PROGRAM PRG_IO_In
VAR
    fbSimInfeed, fbSimOutfeed, fbSimEjector, fbSimClamp, fbSimDiverter : FB_CylinderSim;
    fbSimCW : FB_CwSim;
END_VAR

IF GVL_Ctrl.xSim THEN
    //================ SIMULATION =================
    fbSimInfeed(  xValveWork := GVL_IO.stInfeed.xValveWork,   xValveHome := GVL_IO.stInfeed.xValveHome,
                  xSensWork => GVL_IO.stInfeed.xSensWork,     xSensHome => GVL_IO.stInfeed.xSensHome);
    fbSimOutfeed( xValveWork := GVL_IO.stOutfeed.xValveWork,  xValveHome := GVL_IO.stOutfeed.xValveHome,
                  xSensWork => GVL_IO.stOutfeed.xSensWork,    xSensHome => GVL_IO.stOutfeed.xSensHome);
    fbSimEjector( xValveWork := GVL_IO.stEjector.xValveWork,  xValveHome := GVL_IO.stEjector.xValveHome,
                  xSensWork => GVL_IO.stEjector.xSensWork,    xSensHome => GVL_IO.stEjector.xSensHome);
    fbSimClamp(   xValveWork := GVL_IO.stClamp.xValveWork,    xValveHome := GVL_IO.stClamp.xValveHome,
                  xSensWork => GVL_IO.stClamp.xSensWork,      xSensHome => GVL_IO.stClamp.xSensHome);
    fbSimDiverter(xValveWork := GVL_IO.stDiverter.xValveWork, xValveHome := GVL_IO.stDiverter.xValveHome,
                  xSensWork => GVL_IO.stDiverter.xSensWork,   xSensHome => GVL_IO.stDiverter.xSensHome);

    fbSimCW(xEnable := GVL_IO.xLaserEnable AND GVL_IO.xCW_STO,
            xTrig   := GVL_IO.xCW_Trig,
            nJob    := GVL_IO.nCW_Job,
            xReady  => GVL_IO.xCW_Lready,
            xJobLoaded => GVL_IO.xCW_JobLoaded,
            xBusy   => GVL_IO.xCW_MarkBusy);

    // part leaves the infeed barrier when the infeed cylinder pushed it;
    // part appears at the outfeed barrier after the ejector pushed a GOOD part (no bypass),
    // and disappears when the outfeed cylinder took it.
    IF GVL_IO.stInfeed.xSensWork THEN
        GVL_Ctrl.xSimPartIn := FALSE;
    END_IF
    IF GVL_IO.stEjector.xSensWork AND NOT GVL_IO.xBypassAS THEN
        GVL_Ctrl.xSimPartOut := TRUE;
    ELSIF GVL_IO.stOutfeed.xSensWork THEN
        GVL_Ctrl.xSimPartOut := FALSE;
    END_IF

    GVL_IO.xEStop          := GVL_Ctrl.xSimEStop;
    GVL_IO.xPressureOK     := GVL_Ctrl.xSimPressureOK;
    GVL_IO.xLS_Infeed      := GVL_Ctrl.xSimPartIn;
    GVL_IO.xLS_Outfeed     := GVL_Ctrl.xSimPartOut;
    GVL_IO.xServoInLatched := TRUE;   GVL_IO.xServoInAS  := FALSE;  GVL_IO.xServoInGS  := TRUE;
    GVL_IO.xServoOutLatched:= TRUE;   GVL_IO.xServoOutAS := FALSE;  GVL_IO.xServoOutGS := TRUE;
ELSE
    //================ REAL HARDWARE =================
    GVL_IO.xPressureOK     := GVL_HW.xMaintPressureOK;
    GVL_IO.xEStop          := GVL_HW.xEStopPressed;
    GVL_IO.xLS_Infeed      := GVL_HW.xLS_Infeed;
    GVL_IO.xLS_Outfeed     := GVL_HW.xLS_Outfeed;
    GVL_IO.xServoInLatched := GVL_HW.xServoIn_Latched;
    GVL_IO.xServoInAS      := GVL_HW.xServoIn_AS;
    GVL_IO.xServoInGS      := GVL_HW.xServoIn_GS;
    GVL_IO.xServoOutLatched:= GVL_HW.xServoOut_Latched;
    GVL_IO.xServoOutAS     := GVL_HW.xServoOut_AS;
    GVL_IO.xServoOutGS     := GVL_HW.xServoOut_GS;
    GVL_IO.xCW_Lready      := GVL_HW.xCW_Lready;
    GVL_IO.xCW_JobLoaded   := GVL_HW.xCW_JobLoaded;
    GVL_IO.xCW_MarkBusy    := GVL_HW.xCW_MarkBusy;

    GVL_IO.stInfeed.xSensWork   := GVL_HW.xSnsInfeed_AS;    GVL_IO.stInfeed.xSensHome   := GVL_HW.xSnsInfeed_GS;
    GVL_IO.stOutfeed.xSensWork  := GVL_HW.xSnsOutfeed_AS;   GVL_IO.stOutfeed.xSensHome  := GVL_HW.xSnsOutfeed_GS;
    GVL_IO.stEjector.xSensWork  := GVL_HW.xSnsEjector_AS;   GVL_IO.stEjector.xSensHome  := GVL_HW.xSnsEjector_GS;
    GVL_IO.stClamp.xSensWork    := GVL_HW.xSnsClamp_AS;     GVL_IO.stClamp.xSensHome    := GVL_HW.xSnsClamp_GS;
    GVL_IO.stDiverter.xSensWork := GVL_HW.xSnsDiverter_AS;  GVL_IO.stDiverter.xSensHome := GVL_HW.xSnsDiverter_GS;
END_IF

END_PROGRAM

(* stored: Version 1.1.0.1
   POU PRG_IO_In: Id {94f77fec-ea39-4469-9918-960467030ef8}, SpecialFunc None *)
